KUKA KRL program: ConfProg.src

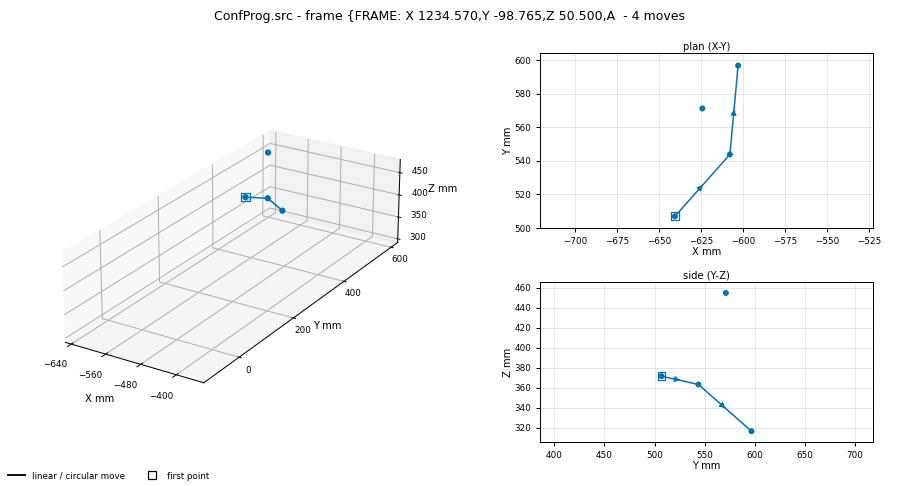
[picture p0: tool path of ConfProg.src in frame {FRAME: X 1234.570,Y -98.765,Z 50.500,A , 4 of 6 moves have a stored position in this frame; points joined in program order, loops and branches not executed]
&ACCESS RVP
&REL 1
&PARAM TEMPLATE = C:\KRC\Roboter\Template\vorgabe
&PARAM EDITMASK = *
DEF ConfProg ( )
EXT BAS (BAS_COMMAND :IN,REAL :IN )


; GLOBAL INTERRUPT DECL 3 WHEN $STOPMESS==TRUE DO IR_STOPM ( )
; INTERRUPT ON 3

;FOLD Initialise and set default speed
BAS (#INITMOV,0)
BAS (#VEL_PTP,100)
BAS (#ACC_PTP,20)
$VEL.CP=0.2
BAS (#TOOL,0)
BAS (#BASE,0)
;ENDFOLD

;;FOLD STARTPOS
;$BWDSTART = FALSE
;PDAT_ACT = PDEFAULT
;BAS(#PTP_DAT)
;FDAT_ACT = {TOOL_NO 0,BASE_NO 0,IPO_FRAME #BASE}
;BAS(#FRAMES)
;;ENDFOLD

$ADVANCE = 5

;FOLD ---- Quickly skip BCO ----
; PTP $AXIS_ACT
;ENDFOLD

;FOLD ---- GO HOME ----
; PTP {A1 0.000, A2 -90.000, A3 90.000, A4 0.000, A5 0.000, A6 0.000, E1 0, E2 0, E3 0, E4 0, E5 0, E6 0}
;ENDFOLD


; Program generated by RoboDK v6.0.7 for KUKA KR 10 R1100-2 on XX/XX/XXXX 18:00:00
; Using nominal kinematics.
; ---- Setting reference (Base) ----
$BASE = {FRAME: X 1234.570,Y -98.765,Z 50.500,A 30.000,B 0.000,C 0.000}
; --------------------------
; ---- Setting tool (TCP) ----
$TOOL = {FRAME: X 10.000,Y 20.000,Z 150.000,A 0.000,B 0.000,C 0.000}
; --------------------------
LIN {X -640.584,Y 506.980,Z 371.534,A 150.000,B 50.000,C -165.000}
LIN {X -607.850,Y 543.849,Z 363.215,A 150.000,B 50.000,C -165.000}
LIN {X -602.951,Y 596.788,Z 316.595,A 150.000,B 50.000,C -165.000}
PTP {A1 10.00000,A2 20.00000,A3 -30.00000,A4 40.00000,A5 -50.00000,A6 60.00000}
PTP {A1 -170.00000,A2 45.00000,A3 -45.00000,A4 -170.00000,A5 90.00000,A6 -179.00000}
CIRC {X -353.026,Y -90.135,Z 331.702,A 178.023,B 40.650,C -169.444},{X -624.230,Y 571.208,Z 454.620,A -122.815,B 44.567,C -82.711}
END
